// TIA Portal V21 export
// export: Created 2026-11-10T07:35:10.2249941Z, ExportSetting WithDefaults, DisplayName Totally Integrated Automation Portal, DisplayVersion V21 Update 3, DisplayName STEP 7 Professional, DisplayVersion V21 Update 3, DisplayName STEP 7 Safety, DisplayVersion V21, DisplayName Tech WebApplication, DisplayVersion V21, DisplayName WinCC Basic/Comfort/Advanced, DisplayVersion V21 Update 3, DisplayName WinCC Unified, DisplayVersion V21 Update 3
FUNCTION_BLOCK "FB_Lad_ex096"   // FB99, LAD
{ S7_Optimized_Access := 'TRUE' }
VERSION : 0.1
// stored: AutoNumber true, IsIECCheckEnabled false, IsRetainMemResEnabled false, MemoryReserve 100, SetENOAutomatically false, UDAEnableTagReadback false
   VAR_INPUT
      v_req : Bool;
      v_laddr : HW_IO;
      v_index : Int;
   END_VAR
   VAR_OUTPUT
      v_valid : Bool;
      v_busy : Bool;
      v_error : Bool;
      v_status : DWord;
      v_len : Int;
   END_VAR
   VAR_IN_OUT
      v_record : Array[0..99] of Byte;
   END_VAR
   VAR
      inst { S7_SetPoint := 'True'} : RD_DPAR;
   END_VAR
BEGIN

REGION Network 1: RD_DPAR - Read module data record
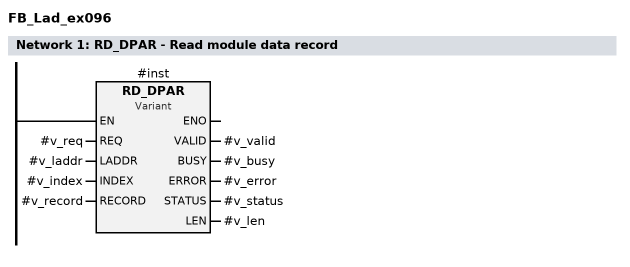
   RUNG wire#powerrail
      { S7_Templates := "[ptr_type := Variant, laddr_type := HW_IO]" } #inst.RD_DPAR(REQ := #v_req, LADDR := #v_laddr, INDEX := #v_index, RECORD := #v_record, VALID => #v_valid, BUSY => #v_busy, ERROR => #v_error, STATUS => #v_status, LEN => #v_len)
   END_RUNG
   // the same network as SCL:
   #inst(REQ := #v_req,   // RD_DPAR
         LADDR := #v_laddr,
         INDEX := #v_index,
         RECORD := #v_record,
         VALID => #v_valid,
         BUSY => #v_busy,
         ERROR => #v_error,
         STATUS => #v_status,
         LEN => #v_len);
END_REGION
END_FUNCTION_BLOCK
